// TIA Portal V20 export
// export: Created 2026-10-12T05:35:23.88251Z, ExportSetting WithDefaults, DisplayName Totally Integrated Automation Portal, DisplayVersion V20, DisplayName TIA Portal Openness, DisplayVersion V20, DisplayName TIA Portal Teamcenter Gateway, DisplayVersion V20, DisplayName TIA Portal Version Control Interface, DisplayVersion V20, DisplayName SINAMICS Startdrive Advanced, DisplayVersion V20 SP1 Update 2, DisplayName SINAMICS Startdrive G110M, G120, G120C, G120D, G120P, G115D, DisplayVersion V20 SP1 Update 2, DisplayName SINAMICS Startdrive G130, G150, S120, S150, SINAMICS MV, G220, S200, S210, DisplayVersion V20 SP1 Update 2, DisplayName STEP 7 Professional, DisplayVersion V20, DisplayName STEP 7 Safety, DisplayVersion V20, DisplayName WinCC Basic/Comfort/Advanced, DisplayVersion V20, DisplayName WinCC Professional, DisplayVersion V20, DisplayName WinCC Unified, DisplayVersion V20
FUNCTION "FRK_AccessCrcByte" : DWord   // FC49, SCL
{ S7_Optimized_Access := 'TRUE' }
VERSION : 0.1
// Reference-1500 LOCAL_RETAIN adapter. No sessions or plaintext credentials.
//  CRC-32 arithmetic comes from Core F_Crc32; encoding is binding-local, versioned.
// stored: AutoNumber true, IsIECCheckEnabled false, SetENOAutomatically false, UDAEnableTagReadback false
   VAR_INPUT
      Previous : DWord;
      Value : Byte;
   END_VAR
   VAR_TEMP
      BitIndex : Int;
      Work : DWord;
   END_VAR
BEGIN

   #Work := #Previous XOR BYTE_TO_DWORD(#Value);
   FOR #BitIndex := 0 TO 7 DO
       IF (#Work AND DWORD#1) <> 0 THEN
           #Work := SHR(IN := #Work, N := 1) XOR DWORD#16#EDB88320;
       ELSE
           #Work := SHR(IN := #Work, N := 1);
       END_IF;
   END_FOR;
   #FRK_AccessCrcByte := #Work;
END_FUNCTION
